// TIA Portal project "038_comm_hw" (V21)

(* hardware
DEVICE "PLC_1"  S7-1500 station
   slot 0: "Rail_0"  Rack  6ES7 590-1***0-0AA0
   slot 1: "PLC_1"  CPU 1513-1 PN  6ES7 513-1AL02-0AB0  V2.9
      slot 3: "CPU display_1"  6ES7591-1AA00-0AA0
      slot 32768: "PROFINET interface_1"  X1
         slot 32769: "Port_1"  X1 P1
         slot 32770: "Port_2"  X1 P2
      slot 34817: "Virtual CP interface port_1"  Virtual CP interface port  Virtual CP interface port
   slot 2: "CM_PtP_1"  CM PtP RS422/485 HF  6ES7 541-1AB00-0AB0  V1.0
*)

// ===== PLC "PLC_1"  CPU 1513-1 PN =====

FUNCTION_BLOCK "FB_Lad_pt006"   // FB1, LAD
{ S7_Optimized_Access := 'TRUE' }
   VAR_INPUT
      v_req : Bool;
      v_port : Port;
   END_VAR
   VAR_OUTPUT
      v_done : Bool;
      v_error : Bool;
      v_status : Word;
   END_VAR
   VAR
      inst : Receive_Reset;
   END_VAR
BEGIN

REGION Network 1: RCV_RST - Delete receive buffer
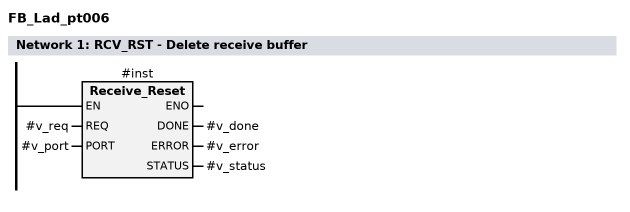
   #inst(REQ := #v_req, PORT := #v_port, DONE => #v_done, ERROR => #v_error, STATUS => #v_status);   // Receive_Reset
END_REGION
END_FUNCTION_BLOCK

FUNCTION_BLOCK "FB_Lad_pt007"   // FB2, LAD
{ S7_Optimized_Access := 'TRUE' }
   VAR_INPUT
      v_req : Bool;
      v_port : Port;
   END_VAR
   VAR_OUTPUT
      v_ndr : Bool;
      v_dtr : Bool;
      v_dsr : Bool;
      v_rts : Bool;
      v_cts : Bool;
      v_dcd : Bool;
      v_ring : Bool;
      v_error : Bool;
      v_status : Word;
   END_VAR
   VAR
      inst : Signal_Get;
   END_VAR
BEGIN

REGION Network 1: SGN_GET - Query RS-232 signals
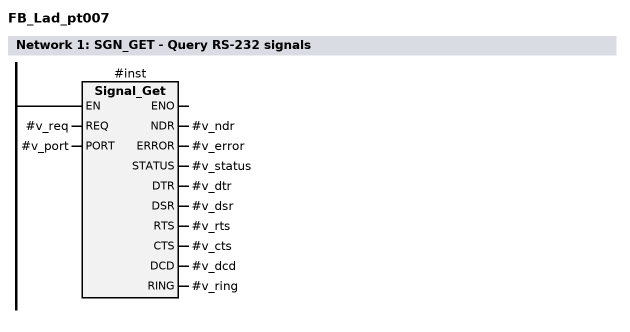
   #inst(REQ := #v_req,   // Signal_Get
         PORT := #v_port,
         NDR => #v_ndr,
         ERROR => #v_error,
         STATUS => #v_status,
         DTR => #v_dtr,
         DSR => #v_dsr,
         RTS => #v_rts,
         CTS => #v_cts,
         DCD => #v_dcd,
         RING => #v_ring);
END_REGION
END_FUNCTION_BLOCK

FUNCTION_BLOCK "FB_Lad_pt008"   // FB3, LAD
{ S7_Optimized_Access := 'TRUE' }
   VAR_INPUT
      v_req : Bool;
      v_port : Port;
      v_signal : Byte;
      v_rts : Bool;
      v_dtr : Bool;
      v_dsr : Bool;
   END_VAR
   VAR_OUTPUT
      v_done : Bool;
      v_error : Bool;
      v_status : Word;
   END_VAR
   VAR
      inst : Signal_Set;
   END_VAR
BEGIN

REGION Network 1: SGN_SET - Set RS-232 signals
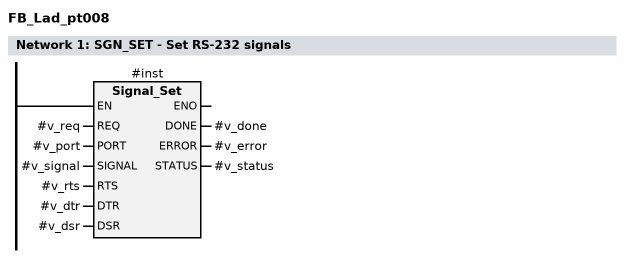
   #inst(REQ := #v_req,   // Signal_Set
         PORT := #v_port,
         SIGNAL := #v_signal,
         RTS := #v_rts,
         DTR := #v_dtr,
         DSR := #v_dsr,
         DONE => #v_done,
         ERROR => #v_error,
         STATUS => #v_status);
END_REGION
END_FUNCTION_BLOCK

FUNCTION_BLOCK "FB_Lad_us004"   // FB4, LAD
{ S7_Optimized_Access := 'TRUE' }
   VAR_INPUT
      v_run : Bool;
      v_off2 : Bool;
      v_off3 : Bool;
      v_f_ack : Bool;
      v_dir : Bool;
      v_drive : USInt;
      v_pzd_len : USInt;
      v_speed_sp : Real;
      v_ctrl3 : Word;
      v_ctrl4 : Word;
      v_ctrl5 : Word;
      v_ctrl6 : Word;
      v_ctrl7 : Word;
      v_ctrl8 : Word;
   END_VAR
   VAR_OUTPUT
      v_ndr : Bool;
      v_error : Bool;
      v_status : Word;
      v_run_en : Bool;
      v_d_dir : Bool;
      v_inhibit : Bool;
      v_fault : Bool;
      v_speed : Real;
      v_status1 : Word;
      v_status3 : Word;
      v_status4 : Word;
      v_status5 : Word;
      v_status6 : Word;
      v_status7 : Word;
      v_status8 : Word;
   END_VAR
   VAR
      inst : USS_Drive_Control;
   END_VAR
BEGIN

REGION Network 1: USS_DRIVE - Swap data with drive
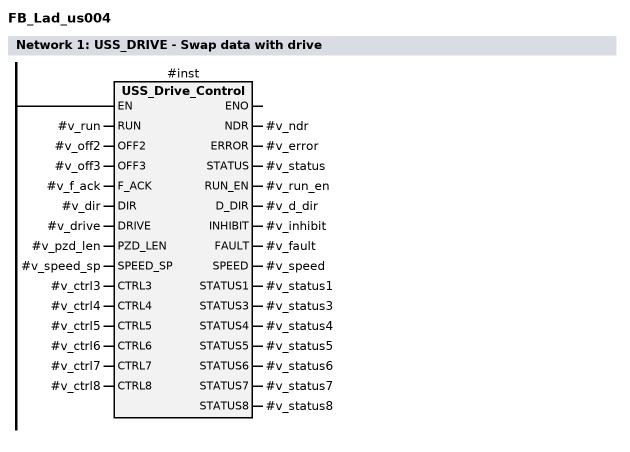
   #inst(RUN := #v_run,   // USS_Drive_Control
         OFF2 := #v_off2,
         OFF3 := #v_off3,
         F_ACK := #v_f_ack,
         DIR := #v_dir,
         DRIVE := #v_drive,
         PZD_LEN := #v_pzd_len,
         SPEED_SP := #v_speed_sp,
         CTRL3 := #v_ctrl3,
         CTRL4 := #v_ctrl4,
         CTRL5 := #v_ctrl5,
         CTRL6 := #v_ctrl6,
         CTRL7 := #v_ctrl7,
         CTRL8 := #v_ctrl8,
         NDR => #v_ndr,
         ERROR => #v_error,
         STATUS => #v_status,
         RUN_EN => #v_run_en,
         D_DIR => #v_d_dir,
         INHIBIT => #v_inhibit,
         FAULT => #v_fault,
         SPEED => #v_speed,
         STATUS1 => #v_status1,
         STATUS3 => #v_status3,
         STATUS4 => #v_status4,
         STATUS5 => #v_status5,
         STATUS6 => #v_status6,
         STATUS7 => #v_status7,
         STATUS8 => #v_status8);
END_REGION
END_FUNCTION_BLOCK

FUNCTION_BLOCK "FB_Lad_mb001"   // FB5, LAD
{ S7_Optimized_Access := 'TRUE' }
   VAR_INPUT
      v_req : Bool;
      v_port : Port;
      v_baud : UDInt;
      v_parity : UInt;
      v_flow_ctrl : UInt;
      v_rts_on_dly : UInt;
      v_rts_off_dly : UInt;
      v_resp_to : UInt;
   END_VAR
   VAR_OUTPUT
      v_done : Bool;
      v_error : Bool;
      v_status : Word;
   END_VAR
   VAR_IN_OUT
      v_mb_db : P2P_MB_BASE;
   END_VAR
   VAR
      inst : Modbus_Comm_Load;
   END_VAR
BEGIN

REGION Network 1: MB_COMM_LOAD - Configure port on the PtP module for Modbus RTU
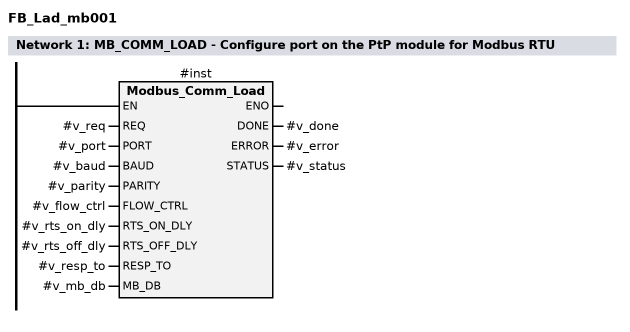
   #inst(REQ := #v_req,   // Modbus_Comm_Load
         PORT := #v_port,
         BAUD := #v_baud,
         PARITY := #v_parity,
         FLOW_CTRL := #v_flow_ctrl,
         RTS_ON_DLY := #v_rts_on_dly,
         RTS_OFF_DLY := #v_rts_off_dly,
         RESP_TO := #v_resp_to,
         MB_DB := #v_mb_db,
         DONE => #v_done,
         ERROR => #v_error,
         STATUS => #v_status);
END_REGION
END_FUNCTION_BLOCK

FUNCTION_BLOCK "FB_Lad_us003"   // FB6, LAD
{ S7_Optimized_Access := 'TRUE' }
   VAR_INPUT
      v_port : Port;
      v_baud : DInt;
   END_VAR
   VAR_OUTPUT
      v_error : Bool;
      v_status : Word;
   END_VAR
   VAR_IN_OUT
      v_uss_db : P2P_USS_BASE;
   END_VAR
   VAR
      inst : USS_Port_Scan;
   END_VAR
BEGIN

REGION Network 1: USS_PORT - Edit communication via USS network
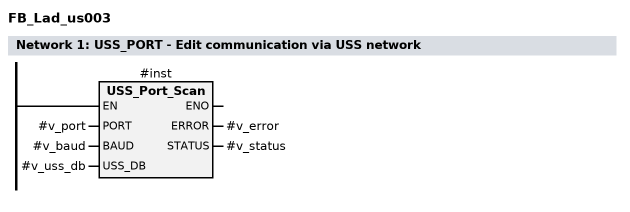
   #inst(PORT := #v_port, BAUD := #v_baud, USS_DB := #v_uss_db, ERROR => #v_error, STATUS => #v_status);   // USS_Port_Scan
END_REGION
END_FUNCTION_BLOCK

FUNCTION_BLOCK "FB_Lad_mb002"   // FB7, LAD
{ S7_Optimized_Access := 'TRUE' }
   VAR_INPUT
      v_req : Bool;
      v_mb_addr : UInt;
      v_mode : USInt;
      v_data_addr : UDInt;
      v_data_len : UInt;
   END_VAR
   VAR_OUTPUT
      v_done : Bool;
      v_busy : Bool;
      v_error : Bool;
      v_status : Word;
   END_VAR
   VAR_IN_OUT
      v_data_ptr : Variant;
   END_VAR
   VAR
      inst : Modbus_Master;
   END_VAR
BEGIN

REGION Network 1: Description of MB_MASTER
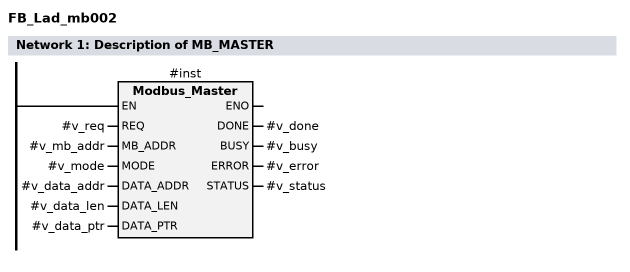
   #inst(REQ := #v_req,   // Modbus_Master
         MB_ADDR := #v_mb_addr,
         MODE := #v_mode,
         DATA_ADDR := #v_data_addr,
         DATA_LEN := #v_data_len,
         DATA_PTR := #v_data_ptr,
         DONE => #v_done,
         BUSY => #v_busy,
         ERROR => #v_error,
         STATUS => #v_status);
END_REGION
END_FUNCTION_BLOCK

FUNCTION_BLOCK "FB_Lad_mb008"   // FB8, LAD
{ S7_Optimized_Access := 'TRUE' }
   VAR_INPUT
      v_mb_addr : USInt;
   END_VAR
   VAR_OUTPUT
      v_ndr : Bool;
      v_dr : Bool;
      v_error : Bool;
      v_status : Word;
   END_VAR
   VAR_IN_OUT
      v_mb_hold_reg : Variant;
   END_VAR
   VAR
      inst : Modbus_Slave;
   END_VAR
BEGIN

REGION Network 1: Description of MB_SLAVE
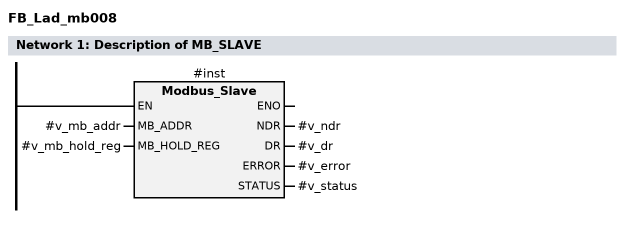
   #inst(MB_ADDR := #v_mb_addr,   // Modbus_Slave
         MB_HOLD_REG := #v_mb_hold_reg,
         NDR => #v_ndr,
         DR => #v_dr,
         ERROR => #v_error,
         STATUS => #v_status);
END_REGION
END_FUNCTION_BLOCK

FUNCTION_BLOCK "FB_Lad_us005"   // FB9, LAD
{ S7_Optimized_Access := 'TRUE' }
   VAR_INPUT
      v_req : Bool;
      v_drive : USInt;
      v_param : UInt;
      v_index : UInt;
   END_VAR
   VAR_OUTPUT
      v_done : Bool;
      v_error : Bool;
      v_status : Word;
   END_VAR
   VAR_IN_OUT
      v_uss_db : P2P_USS_BASE;
      v_value : P2P_USS_BASE;
   END_VAR
BEGIN

REGION Network 1: USS_RPM - Readout parameters from the drive
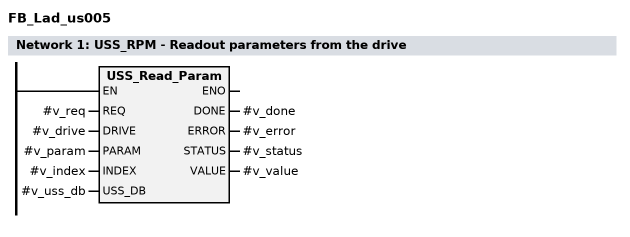
   // no SCL statement known for USS_Read_Param: written as a call
   USS_Read_Param(REQ := #v_req,
                  DRIVE := #v_drive,
                  PARAM := #v_param,
                  INDEX := #v_index,
                  USS_DB := #v_uss_db,
                  DONE => #v_done,
                  ERROR => #v_error,
                  STATUS => #v_status,
                  VALUE => #v_value);
END_REGION
END_FUNCTION_BLOCK

FUNCTION_BLOCK "FB_Lad_us006"   // FB10, LAD
{ S7_Optimized_Access := 'TRUE' }
   VAR_INPUT
      v_req : Bool;
      v_drive : USInt;
      v_param : UInt;
      v_index : UInt;
      v_eeprom : Bool;
      v_value : P2P_USS_BASE;
   END_VAR
   VAR_OUTPUT
      v_done : Bool;
      v_error : Bool;
      v_status : Word;
   END_VAR
   VAR_IN_OUT
      v_uss_db : P2P_USS_BASE;
   END_VAR
BEGIN

REGION Network 1: USS_WPM - Change parameters in the drive
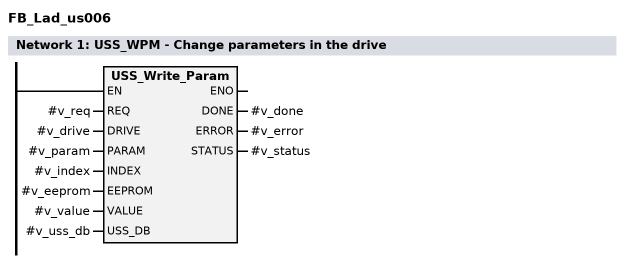
   // no SCL statement known for USS_Write_Param: written as a call
   USS_Write_Param(REQ := #v_req,
                   DRIVE := #v_drive,
                   PARAM := #v_param,
                   INDEX := #v_index,
                   EEPROM := #v_eeprom,
                   VALUE := #v_value,
                   USS_DB := #v_uss_db,
                   DONE => #v_done,
                   ERROR => #v_error,
                   STATUS => #v_status);
END_REGION
END_FUNCTION_BLOCK

ORGANIZATION_BLOCK "Main"   // OB1, LAD, ProgramCycle
TITLE = "Main Program Sweep (Cycle)"
{ S7_Optimized_Access := 'TRUE' }
VERSION : 0.1
   VAR_INPUT
      Initial_Call : Bool;   // Initial call of this OB
      Remanence : Bool;   // =True, if remanent data are available
   END_VAR
BEGIN
END_ORGANIZATION_BLOCK